Fanuc KAREL source: KT00737.KL

PROGRAM KT00737
%NOLOCKGROUP
VAR
  ARG: ARRAY[4] OF STRING[20]
  OUT: INTEGER
BEGIN
  OUT = ARRAY_LEN(ARG)
END KT00737
